// TIA Portal V19 export
FUNCTION_BLOCK "RAMP"   // FB12, LAD
{ S7_Optimized_Access := 'TRUE' }
// stored: MemoryReserve 100, SetENOAutomatically false
   VAR_INPUT
      RAMP_START : Bool;
      JACKET_TT02 : Real;
      MASS_TT03 : Real;
      PRODUCT_TT : Real;
      RESET : Bool;
      SP : Real;
      PV : Real;
      "TIME" : Int;
      MAIN_START : Bool;
      MAIN_TIME : Int;
      MAIN_RESET : Bool;
      JACKET : Bool;
      MASS : Bool;
      PRODUCT : Bool;
      "A/M" : Bool;
      TIMER_RESET : Bool;
      COOL_RUNNING : Bool;
      HEAT_RUUNNING : Bool;
      SEMI : Bool;
   END_VAR
   VAR_OUTPUT
      RAMP_SP : Real;
      RAMP_RATE : Real;
      MAIN_COM : Bool;
      MAIN_PV : Real;
      RAMP_MIN : Int;
   END_VAR
   VAR_IN_OUT
      RAMP_INPUT : Real;
      TIME_1 : Int;
      ramp_substitute : Real;
   END_VAR
   VAR
      RampFunction_Instance { S7_SetPoint := 'True'} : RampFunction;
      TIMER_SECONDS_Instance { S7_SetPoint := 'True'} : "TIMER_SECONDS";
      START_MAIN_TIMER { S7_SetPoint := 'True'} : Bool;
      RAMP_TEMP_OUT : Real;
      TIMER_SECONDS_Instance_1 { S7_SetPoint := 'True'} : "TIMER_SECONDS";
      RAMP_CV_CTL { S7_SetPoint := 'True'} : PID_Compact;
      PID_Compact_1 { S7_SetPoint := 'True'} : PID_Compact;
      NORM_MIN : Int;
      NORM_MAX : Int;
      SCALE_MIN : Real;
      SCALE_MAX : Real;
      MAN_INPUT : Int;
      NORM_OUT : Real;
      SCVOUT : Int;
      MANOUT : Int;
      AO : Int;
      TIMER_SECONDS_Instance_2 { S7_SetPoint := 'True'} : "TIMER_SECONDS";
      P_TRIG6 { S7_SetPoint := 'True'} : Bool;
      P_TRIG7 : Bool;
      SEC : Int;
      IEC_Timer_0_Instance { S7_SetPoint := 'True'} : TOF_TIME;
      IEC_Timer_0_Instance_1 { S7_SetPoint := 'True'} : TP_TIME;
   END_VAR
   // RAMP_CV_CTL.Mode := 2;
   // RAMP_CV_CTL.PhysicalQuantity := 1;
   // RAMP_CV_CTL.Config.InputPerOn := FALSE;
   // RAMP_CV_CTL.Config.InputUpperLimit := 200.0;
   VAR_TEMP   // added for the SCL form of the ladder/FBD networks
      _w1 : Bool;
      _w2 : Bool;
      _w3 : Bool;
      _w4 : Bool;
   END_VAR
BEGIN

REGION Network 1
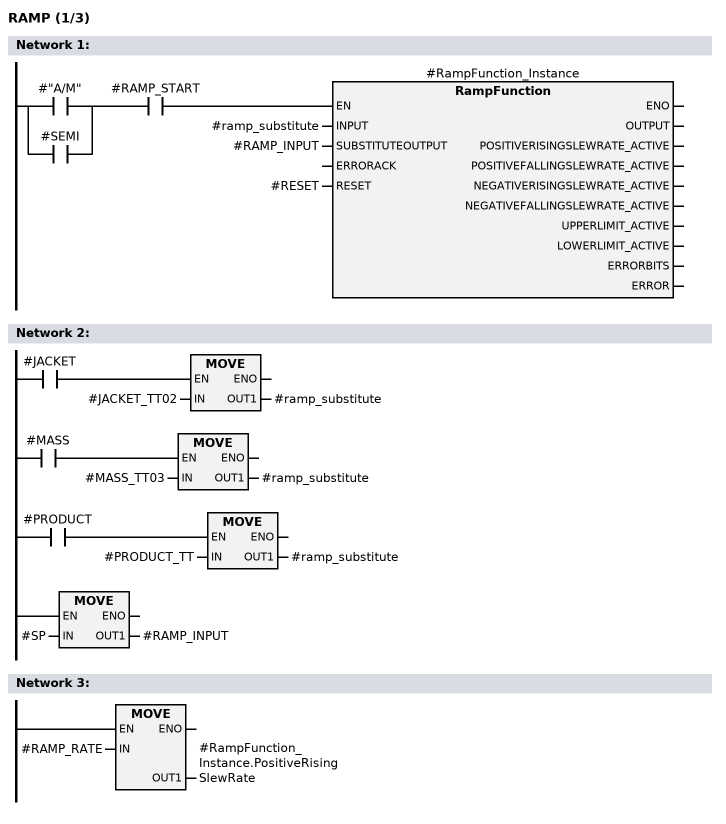
   RUNG wire#powerrail
      Contact( #"A/M" )
      wire#w1
      Contact( #RAMP_START )
      #RampFunction_Instance.RampFunction(Input := #ramp_substitute, SubstituteOutput := #RAMP_INPUT, ErrorAck :=, Reset := #RESET, Output =>, PositiveRisingSlewRate_Active =>, PositiveFallingSlewRate_Active =>, NegativeRisingSlewRate_Active =>, NegativeFallingSlewRate_Active =>, UpperLimit_Active =>, LowerLimit_Active =>, ErrorBits =>, Error =>)
   END_RUNG
   RUNG wire#powerrail
      Contact( #SEMI )
   END_RUNG wire#w1
   // the same network as SCL:
   IF (#"A/M" OR #SEMI) AND #RAMP_START THEN
       #RampFunction_Instance(Input := #ramp_substitute, SubstituteOutput := #RAMP_INPUT, Reset := #RESET);   // RampFunction
   END_IF;
END_REGION

REGION Network 2
   RUNG wire#powerrail
      Contact( #JACKET )
      Move(in := #JACKET_TT02, out1 => #ramp_substitute)
   END_RUNG
   RUNG wire#powerrail
      Contact( #MASS )
      Move(in := #MASS_TT03, out1 => #ramp_substitute)
   END_RUNG
   RUNG wire#powerrail
      Contact( #PRODUCT )
      Move(in := #PRODUCT_TT, out1 => #ramp_substitute)
   END_RUNG
   RUNG wire#powerrail
      Move(in := #SP, out1 => #RAMP_INPUT)
   END_RUNG
   // the same network as SCL:
   IF #JACKET THEN #ramp_substitute := #JACKET_TT02; END_IF;
   IF #MASS THEN #ramp_substitute := #MASS_TT03; END_IF;
   IF #PRODUCT THEN #ramp_substitute := #PRODUCT_TT; END_IF;
   #RAMP_INPUT := #SP;
END_REGION

REGION Network 3
   RUNG wire#powerrail
      Move(in := #RAMP_RATE, out1 => #RampFunction_Instance.PositiveRisingSlewRate)
   END_RUNG
   // the same network as SCL:
   #RampFunction_Instance.PositiveRisingSlewRate := #RAMP_RATE;
END_REGION

REGION Network 4
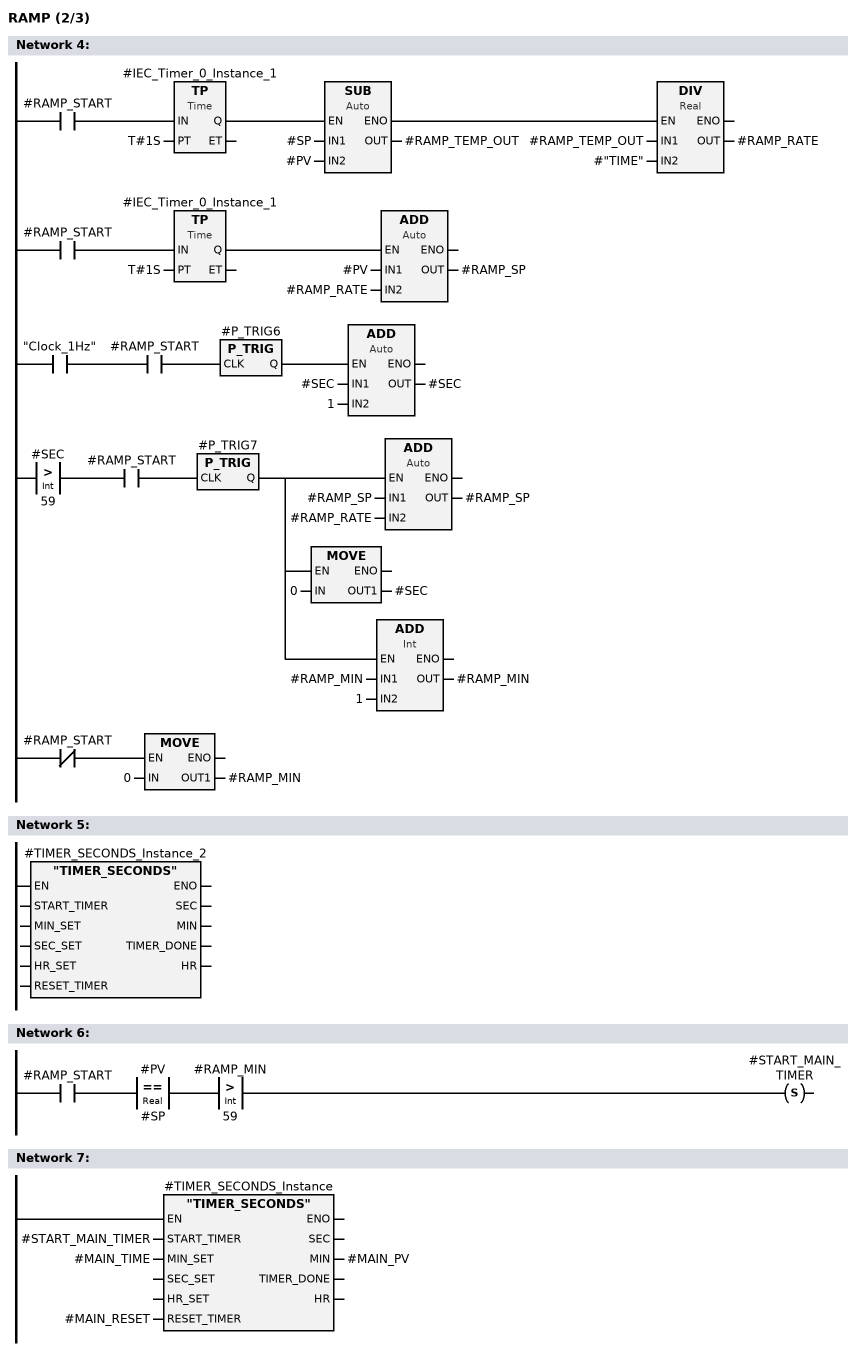
   RUNG wire#powerrail
      Contact( #RAMP_START )
      { S7_Templates := "time_type := Time" } #IEC_Timer_0_Instance_1.TP(pt := T#1S, et =>)
      Sub(in1 := #SP, in2 := #PV, out => #RAMP_TEMP_OUT)
      { S7_Templates := "SrcType := Real" } Div(in1 := #RAMP_TEMP_OUT, in2 := #"TIME", out => #RAMP_RATE)
   END_RUNG
   RUNG wire#powerrail
      Contact( #RAMP_START )
      { S7_Templates := "time_type := Time" } #IEC_Timer_0_Instance_1.TP(pt := T#1S, et =>)
      Add(in1 := #PV, in2 := #RAMP_RATE, out => #RAMP_SP)
   END_RUNG
   RUNG wire#powerrail
      Contact( "Clock_1Hz" )
      Contact( #RAMP_START )
      P_Trig( #P_TRIG6 )
      Add(in1 := #SEC, in2 := 1, out => #SEC)
   END_RUNG
   RUNG wire#powerrail
      { S7_Templates := "SrcType := Int" } GT_Contact(in1 := #SEC, in2 := 59)
      Contact( #RAMP_START )
      P_Trig( #P_TRIG7 )
      wire#w1
      Add(in1 := #RAMP_SP, in2 := #RAMP_RATE, out => #RAMP_SP)
   END_RUNG
   RUNG wire#w1
      Move(in := 0, out1 => #SEC)
   END_RUNG
   RUNG wire#w1
      { S7_Templates := "SrcType := Int" } Add(in1 := #RAMP_MIN, in2 := 1, out => #RAMP_MIN)
   END_RUNG
   RUNG wire#powerrail
      I_Contact( #RAMP_START )
      Move(in := 0, out1 => #RAMP_MIN)
   END_RUNG
   // the same network as SCL:
   #IEC_Timer_0_Instance_1(IN := #RAMP_START, PT := T#1S);   // TP
   IF #IEC_Timer_0_Instance_1.Q THEN
       #RAMP_TEMP_OUT := #SP - #PV;
       #RAMP_RATE := #RAMP_TEMP_OUT / #"TIME";
   END_IF;
   #IEC_Timer_0_Instance_1(IN := #RAMP_START, PT := T#1S);   // TP
   IF #IEC_Timer_0_Instance_1.Q THEN #RAMP_SP := #PV + #RAMP_RATE; END_IF;
   #_w1 := "Clock_1Hz" AND #RAMP_START;
   #_w2 := #_w1 AND NOT #P_TRIG6;   // rising edge
   #P_TRIG6 := #_w1;
   IF #_w2 THEN #SEC := #SEC + 1; END_IF;
   #_w3 := (#SEC > 59) AND #RAMP_START;
   #_w4 := #_w3 AND NOT #P_TRIG7;   // rising edge
   #P_TRIG7 := #_w3;
   IF #_w4 THEN
       #RAMP_SP := #RAMP_SP + #RAMP_RATE;
       #SEC := 0;
       #RAMP_MIN := #RAMP_MIN + 1;
   END_IF;
   IF NOT #RAMP_START THEN #RAMP_MIN := 0; END_IF;
END_REGION

REGION Network 5
   RUNG wire#powerrail
      #TIMER_SECONDS_Instance_2(START_TIMER :=, MIN_SET :=, SEC_SET :=, HR_SET :=, RESET_TIMER :=, SEC =>, MIN =>, TIMER_DONE =>, HR =>)
   END_RUNG
   // the same network as SCL:
   #TIMER_SECONDS_Instance_2();   // "TIMER_SECONDS"
END_REGION

REGION Network 6
   RUNG wire#powerrail
      Contact( #RAMP_START )
      { S7_Templates := "SrcType := Real" } EQ_Contact(in1 := #PV, in2 := #SP)
      { S7_Templates := "SrcType := Int" } GT_Contact(in1 := #RAMP_MIN, in2 := 59)
      S_Coil( #START_MAIN_TIMER )
   END_RUNG
   // the same network as SCL:
   IF #RAMP_START AND (#PV = #SP) AND (#RAMP_MIN > 59) THEN #START_MAIN_TIMER := TRUE; END_IF;
END_REGION

REGION Network 7
   RUNG wire#powerrail
      #TIMER_SECONDS_Instance(START_TIMER := #START_MAIN_TIMER, MIN_SET := #MAIN_TIME, SEC_SET :=, HR_SET :=, RESET_TIMER := #MAIN_RESET, SEC =>, MIN => #MAIN_PV, TIMER_DONE =>, HR =>)
   END_RUNG
   // the same network as SCL:
   #TIMER_SECONDS_Instance(START_TIMER := #START_MAIN_TIMER,   // "TIMER_SECONDS"
                           MIN_SET := #MAIN_TIME,
                           RESET_TIMER := #MAIN_RESET,
                           MIN => #MAIN_PV);
END_REGION

REGION Network 8
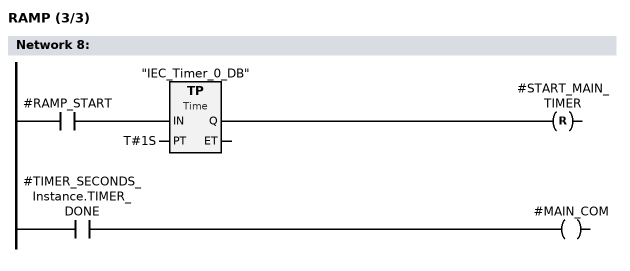
   RUNG wire#powerrail
      Contact( #RAMP_START )
      { S7_Templates := "time_type := Time" } "IEC_Timer_0_DB".TP(pt := T#1S, et =>)
      R_Coil( #START_MAIN_TIMER )
   END_RUNG
   RUNG wire#powerrail
      Contact( #TIMER_SECONDS_Instance.TIMER_DONE )
      Coil( #MAIN_COM )
   END_RUNG
   // the same network as SCL:
   "IEC_Timer_0_DB".TP(IN := #RAMP_START, PT := T#1S);
   IF "IEC_Timer_0_DB".Q THEN #START_MAIN_TIMER := FALSE; END_IF;
   #MAIN_COM := #TIMER_SECONDS_Instance.TIMER_DONE;
END_REGION
END_FUNCTION_BLOCK
